PROGRAM main
  VAR
    S1 AT %IX0.0 : BOOL; (* barrera de entrada: entra un auto *)
    S2 AT %IX0.1 : BOOL; (* barrera de salida: sale un auto *)
    H1 AT %QX0.0 : BOOL; (* verde: hay lugar *)
    H2 AT %QX0.1 : BOOL; (* amarillo: lleno *)
    F_ENTRA      : R_TRIG;
    F_SALE       : R_TRIG;
    AUTOS        : INT; (* autos adentro *)
    LIBRES       : INT; (* lugares libres *)
    ENTRA        : BOOL; (* flanco de S1 *)
    SALE         : BOOL; (* flanco de S2 *)
    HAY_LUGAR    : BOOL; (* AUTOS < capacidad *)
    HAY_AUTOS    : BOOL; (* AUTOS > 0 *)
  END_VAR
  VAR  (* added by the conversion: wires and edge detectors of the diagram *)
    _LT7_OUT : BOOL;
    _GT11_OUT : BOOL;
    _AND16_OUT : BOOL;
    _ADD20_OUT : INT;
    _SEL15_OUT : INT;
    _AND25_OUT : BOOL;
    _SUB29_OUT : INT;
    _SEL24_OUT : INT;
    _SUB33_OUT : INT;
    _GT37_OUT : BOOL;
    _EQ41_OUT : BOOL;
  END_VAR

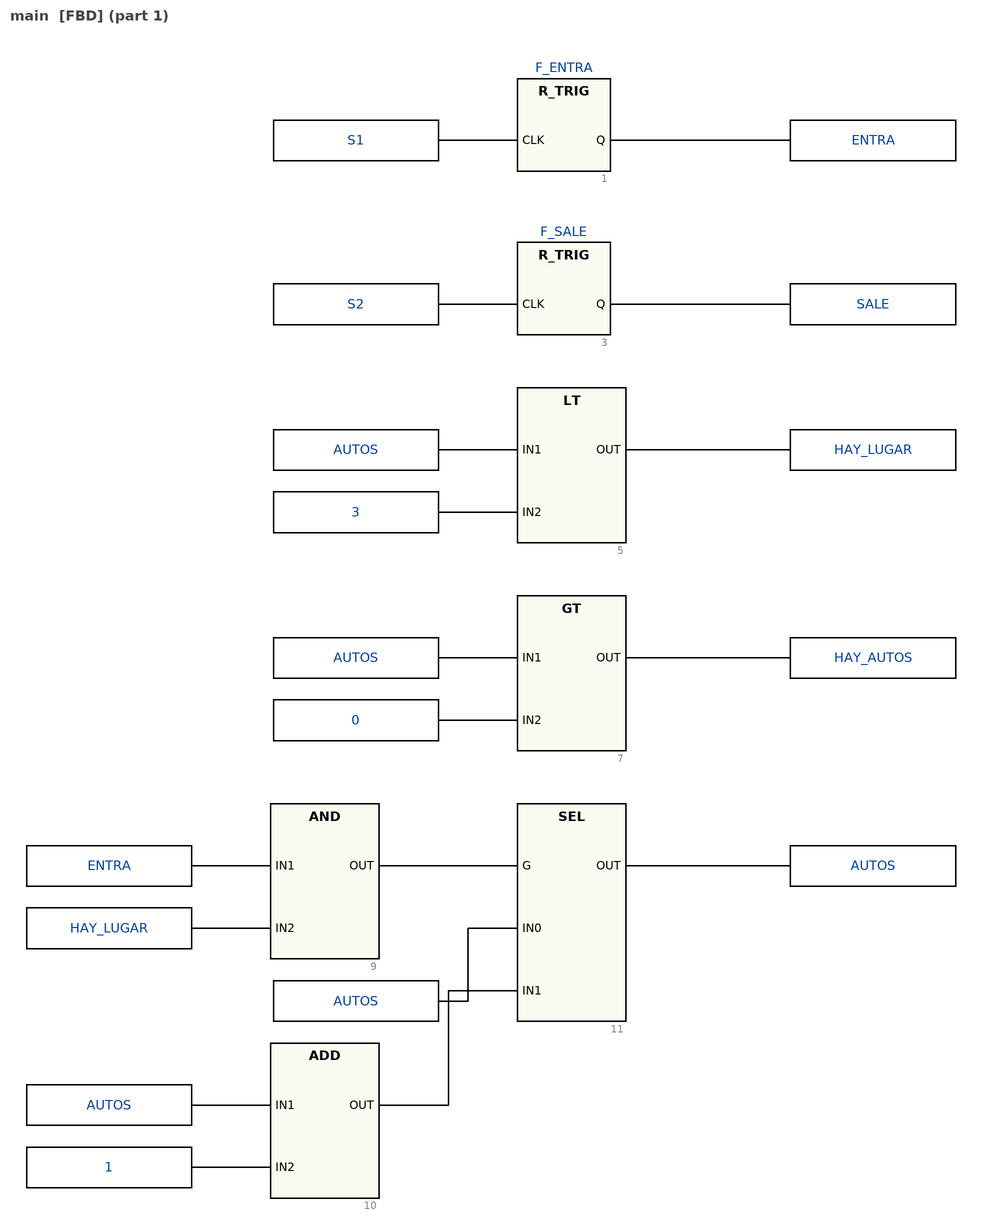
(* FBD diagram, written out as Structured Text *)
F_ENTRA(CLK := S1);
ENTRA := F_ENTRA.Q;
F_SALE(CLK := S2);
SALE := F_SALE.Q;
_LT7_OUT := AUTOS < 3;
HAY_LUGAR := _LT7_OUT;
_GT11_OUT := AUTOS > 0;
HAY_AUTOS := _GT11_OUT;
_AND16_OUT := ENTRA AND HAY_LUGAR;
_ADD20_OUT := AUTOS + 1;
_SEL15_OUT := SEL(_AND16_OUT, AUTOS, _ADD20_OUT);
AUTOS := _SEL15_OUT;
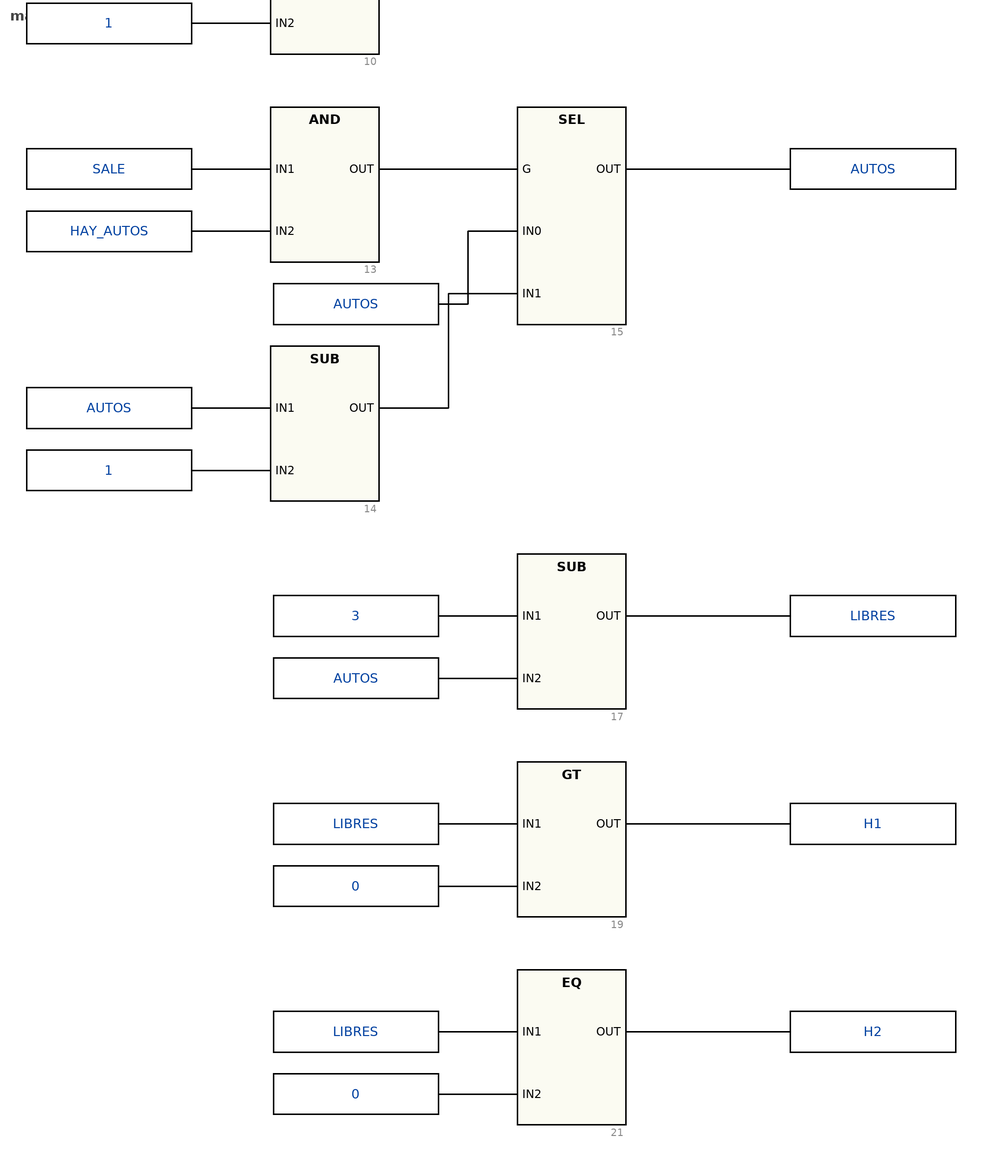
_AND25_OUT := SALE AND HAY_AUTOS;
_SUB29_OUT := AUTOS - 1;
_SEL24_OUT := SEL(_AND25_OUT, AUTOS, _SUB29_OUT);
AUTOS := _SEL24_OUT;
_SUB33_OUT := 3 - AUTOS;
LIBRES := _SUB33_OUT;
_GT37_OUT := LIBRES > 0;
H1 := _GT37_OUT;
_EQ41_OUT := LIBRES = 0;
H2 := _EQ41_OUT;
END_PROGRAM
